(* PLC project coils, tcpethernet coils 1 *)
(* stored: creationDateTime 2026-10-28T09:00:00, modificationDateTime 2026-10-28T09:00:00 *)

PROGRAM coils
  VAR
    A AT %IX0.4 : BOOL;
    B AT %IX0.5 : BOOL;
  END_VAR
  VAR
    Latched : BOOL;
    Edges : INT;
    Pulsed : BOOL;
    Fell : BOOL;
  END_VAR
  VAR  (* added by the conversion: wires and edge detectors of the diagram *)
    R_TRIG1 : R_TRIG;
    _ADD9_ENO : BOOL;
    _ADD9_OUT : INT;
    F_TRIG2 : F_TRIG;
  END_VAR

(* LD diagram, written out as Structured Text *)
IF A THEN Latched := TRUE; END_IF;
IF B THEN Latched := FALSE; END_IF;
R_TRIG1(CLK := A);
_ADD9_OUT := ADD(EN := R_TRIG1.Q, IN1 := Edges, IN2 := 1, ENO => _ADD9_ENO);
Pulsed := _ADD9_ENO;
IF _ADD9_ENO THEN Edges := _ADD9_OUT; END_IF;
F_TRIG2(CLK := A);
Fell := F_TRIG2.Q;
END_PROGRAM
